INTERFACE I_CoverState

METHOD CloseCommand : BOOL
VAR_INPUT
END_VAR
END_METHOD

METHOD OpenCommand : BOOL
VAR_INPUT
END_VAR
END_METHOD

METHOD RunState : BOOL
VAR_INPUT
END_VAR
END_METHOD

METHOD StopCommand : BOOL
VAR_INPUT
END_VAR
END_METHOD

METHOD SuccessfulFinished : BOOL
VAR_INPUT
END_VAR
END_METHOD

END_INTERFACE

(* stored: Version 1.1.0.1, ProductVersion 3.1.4024.15
   Itf I_CoverState: Id {c317b290-0871-446b-945b-a87c63a57de9}
   Method CloseCommand: Id {865f94c7-6c92-4892-a6a4-fe0ec6720f64}
   Method OpenCommand: Id {ab3f11be-d9ee-46fd-bda9-a65c1e611ca1}
   Method RunState: Id {4738b1da-e131-4f8a-9dff-6d4bd4b35c2a}
   Method StopCommand: Id {fbe05262-7bd0-49b3-973f-ed2b5ab7a544}
   Method SuccessfulFinished: Id {40b8cd3b-7ebd-4a9a-9ffc-802528f3077b} *)
